FUNCTION_BLOCK EQ_NeedleAxis (* An equipment block: the only block that touches this equipment's pins. Skills send it what to switch over a local channel; it switches the outputs (off first, then on), reads the inputs every cycle and reports them to the skills and to OPC UA. One skill holds it at a time; on release or when the module aborts it switches everything off. Technical: Needle lift with down/up valves, end switches and a position sensor; equipment IO: owns its IO points, writes the output values its holder sends, reads its inputs every cycle and reports changes *)
  (* Standard: 61499-2 *)
  (* Version 0.1, 2026-09-28, Project contributors, AAU Smart Production Lab *)
  PACKAGE filler;
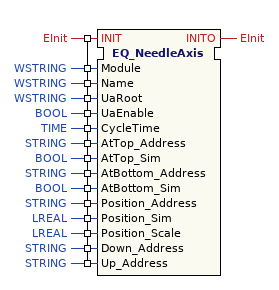
  EVENT_INPUT
    INIT : EInit WITH Module, Name, UaRoot, UaEnable, CycleTime, AtTop_Address, AtTop_Sim, AtBottom_Address, AtBottom_Sim, Position_Address, Position_Sim, Position_Scale, Down_Address, Up_Address; (* Initialise, once at start-up (the INIT chain); takes the values given with it *)
  END_EVENT
  EVENT_OUTPUT
    INITO : EInit; (* Initialised: the next block of the INIT chain goes on *)
  END_EVENT
  VAR_INPUT
    Module : WSTRING; (* The module's name; its local channels are named after it (loc[<Module>/...]) *)
    Name : WSTRING := "NeedleAxis"; (* The equipment item's name: its local channels and OPC UA folder *)
    UaRoot : WSTRING; (* The module's OPC UA folder, e.g. /Objects/Filling *)
    UaEnable : BOOL; (* Publish on OPC UA *)
    CycleTime : TIME := T#50ms; (* How often the inputs are read *)
    AtTop_Address : STRING; (* Where AtTop is: 'gpio[chip:line(:pull_up|:pull_down)(:active_low)]', 'pwm[chip:channel:period_ns]', 'modbus[...]', 'sim', or an IO handle's name; empty: not connected *)
    AtTop_Sim : BOOL := FALSE; (* The value of AtTop when simulated (address 'sim') *)
    AtBottom_Address : STRING; (* Where AtBottom is: 'gpio[chip:line(:pull_up|:pull_down)(:active_low)]', 'pwm[chip:channel:period_ns]', 'modbus[...]', 'sim', or an IO handle's name; empty: not connected *)
    AtBottom_Sim : BOOL := FALSE; (* The value of AtBottom when simulated (address 'sim') *)
    Position_Address : STRING; (* Where Position is: 'gpio[chip:line(:pull_up|:pull_down)(:active_low)]', 'pwm[chip:channel:period_ns]', 'modbus[...]', 'sim', or an IO handle's name; empty: not connected *)
    Position_Sim : LREAL := 0.0; (* The value of Position when simulated (address 'sim') *)
    Position_Scale : LREAL := 0.1; (* Engineering value per raw count of Position *)
    Down_Address : STRING; (* Where Down is: 'gpio[chip:line(:pull_up|:pull_down)(:active_low)]', 'pwm[chip:channel:period_ns]', 'modbus[...]', 'sim', or an IO handle's name; empty: not connected *)
    Up_Address : STRING; (* Where Up is: 'gpio[chip:line(:pull_up|:pull_down)(:active_low)]', 'pwm[chip:channel:period_ns]', 'modbus[...]', 'sim', or an IO handle's name; empty: not connected *)
  END_VAR
  (* Group Core: One holder at a time, break before make, all off on release or abort; scanned every CycleTime *)
  (* Group Channels: Local channels to and from the skills (cmd, release, state), the module's state, and the inputs over OPC UA *)
  (* Group Inputs: The equipment's sensors: read every cycle, one block per IO point *)
  (* Group Outputs: The equipment's actuators: written on a change and every cycle, one block per IO point *)
  FBS
    Logic : filler::EL_NeedleAxis; (* The equipment's logic (EL_): takes commands from one holder at a time, switches the outputs (off first, then on), switches all off on release or module abort, and reports input changes. *) {SET_ATTRIBUTE(GroupName, Core)}
    Cycle : iec61499::events::E_CYCLE; (* Ticks every cycle so the inputs are read and the outputs refreshed. *) {SET_ATTRIBUTE(GroupName, Core)}
    Mode : modlib::MOD_StateView; (* Watches the module's PackML state, to switch everything off when the module aborts. *) {SET_ATTRIBUTE(GroupName, Channels)}
    SubCmd : iec61499::net::SUBSCRIBE_4(QI := TRUE); (* Receives the commands skills send on this equipment's command channel. *) {SET_ATTRIBUTE(GroupName, Channels)}
    SubRelease : iec61499::net::SUBSCRIBE_1(QI := TRUE); (* Hears the module's release channel: when its holder gives up, everything goes off. *) {SET_ATTRIBUTE(GroupName, Channels)}
    PubState : iec61499::net::PUBLISH_4(QI := TRUE); (* Publishes the inputs and the holder on this equipment's state channel, for the skills. *) {SET_ATTRIBUTE(GroupName, Channels)}
    PubUa : iec61499::net::PUBLISH_3; (* Writes the inputs (and a position, if it keeps one) to OPC UA, below Equipment/<item>. *) {SET_ATTRIBUTE(GroupName, Channels)}
    In_AtTop : modlib::IO_DI; (* The pin AtTop: reads the input at AtTop_Address (a Pi pin, Modbus, or simulated). *) {SET_ATTRIBUTE(GroupName, Inputs)}
    In_AtBottom : modlib::IO_DI; (* The pin AtBottom: reads the input at AtBottom_Address (a Pi pin, Modbus, or simulated). *) {SET_ATTRIBUTE(GroupName, Inputs)}
    In_Position : modlib::IO_AI; (* The pin Position: reads the input at Position_Address (a Pi pin, Modbus, or simulated). *) {SET_ATTRIBUTE(GroupName, Inputs)}
    Out_Down : modlib::IO_DO; (* The pin Down: switches the output at Down_Address (a Pi pin, Modbus, or simulated). *) {SET_ATTRIBUTE(GroupName, Outputs)}
    Out_Up : modlib::IO_DO; (* The pin Up: switches the output at Up_Address (a Pi pin, Modbus, or simulated). *) {SET_ATTRIBUTE(GroupName, Outputs)}
  END_FBS
  EVENT_CONNECTIONS
    INIT TO Logic.INIT;
    Logic.INITO TO Mode.INIT;
    Mode.INITO TO SubCmd.INIT;
    SubCmd.INITO TO SubRelease.INIT;
    SubRelease.INITO TO PubState.INIT;
    PubState.INITO TO PubUa.INIT;
    PubUa.INITO TO In_AtTop.INIT;
    In_AtTop.INITO TO In_AtBottom.INIT;
    In_AtBottom.INITO TO In_Position.INIT;
    In_Position.INITO TO Out_Down.INIT;
    Out_Down.INITO TO Out_Up.INIT;
    Out_Up.INITO TO Cycle.START;
    Out_Up.INITO TO INITO;
    SubCmd.IND TO Logic.CMD;
    SubRelease.IND TO Logic.RELEASE;
    Mode.CHG TO Logic.MOD_CHG;
    Cycle.EO TO Logic.REFRESH;
    Cycle.EO TO In_AtTop.REQ;
    In_AtTop.CNF TO In_AtBottom.REQ;
    In_AtBottom.CNF TO In_Position.REQ;
    In_Position.CNF TO Logic.SAMPLE;
    Logic.STATE TO PubState.REQ;
    Logic.STATE TO PubUa.REQ;
    Logic.DRIVE TO Out_Down.REQ;
    Out_Down.CNF TO Out_Up.REQ;
    Out_Up.CNF TO Logic.DRIVEN;
  END_CONNECTIONS
  DATA_CONNECTIONS
    Module TO Logic.Module;
    Name TO Logic.Name;
    UaRoot TO Logic.UaRoot;
    Module TO Mode.Module;
    Logic.IdCmd TO SubCmd.ID;
    Logic.IdRelease TO SubRelease.ID;
    Logic.IdState TO PubState.ID;
    Logic.IdPub TO PubUa.ID;
    UaEnable TO PubUa.QI;
    CycleTime TO Cycle.DT;
    SubCmd.RD_1 TO Logic.C_Holder;
    SubCmd.RD_2 TO Logic.C_Release;
    SubCmd.RD_3 TO Logic.C_Down;
    SubCmd.RD_4 TO Logic.C_Up;
    SubRelease.RD_1 TO Logic.R_Holder;
    Mode.State TO Logic.ModuleState;
    AtTop_Address TO In_AtTop.Address;
    AtTop_Sim TO In_AtTop.SimValue;
    In_AtTop.IN TO Logic.I_AtTop;
    Logic.AtTop TO PubState.SD_1;
    Logic.AtTop TO PubUa.SD_1;
    AtBottom_Address TO In_AtBottom.Address;
    AtBottom_Sim TO In_AtBottom.SimValue;
    In_AtBottom.IN TO Logic.I_AtBottom;
    Logic.AtBottom TO PubState.SD_2;
    Logic.AtBottom TO PubUa.SD_2;
    Position_Address TO In_Position.Address;
    Position_Sim TO In_Position.SimValue;
    Position_Scale TO In_Position.Scale;
    In_Position.IN TO Logic.I_Position;
    Logic.Position TO PubState.SD_3;
    Logic.Position TO PubUa.SD_3;
    Logic.Holder TO PubState.SD_4;
    Down_Address TO Out_Down.Address;
    Logic.O_Down TO Out_Down.OUT;
    Up_Address TO Out_Up.Address;
    Logic.O_Up TO Out_Up.OUT;
  END_CONNECTIONS
END_FUNCTION_BLOCK
